(* PLC project Vn_fb_rs, Beckhoff Automation GmbH TwinCAT PLC Control 3.5.13.21 *)
(* stored: creationDateTime 1970-01-01T00:00:00 *)

PROGRAM Vn_fb_rs

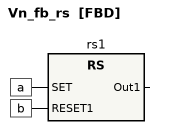
(* FBD diagram, written out as Structured Text *)
rs1(SET := a, RESET1 := b);
END_PROGRAM
